FUNCTION_BLOCK StartStopEvent (* Basic Function Block Type *)
  (* Standard: 61499-2 *)
  (* Version 0.0, 10/21/2026, Schneider Electric, Template *)
  PACKAGE SE.Nereda;
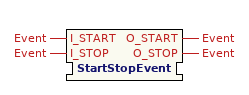
  EVENT_INPUT
    I_START; (* Normal Execution Request *)
    I_STOP;
  END_EVENT
  EVENT_OUTPUT
    O_START; (* Execution Confirmation *)
    O_STOP; (* Initialization Confirm *)
  END_EVENT
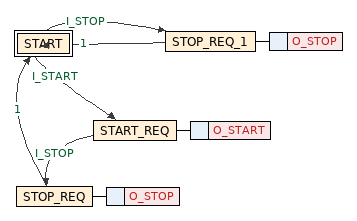
  EC_STATES
    START; (* Initial State *)
    START_REQ : -> O_START;
    STOP_REQ : -> O_STOP;
    STOP_REQ_1 : -> O_STOP;
  END_STATES
  EC_TRANSITIONS
    START TO START_REQ := I_START;
    START_REQ TO STOP_REQ := I_STOP;
    STOP_REQ TO START := 1;
    START TO STOP_REQ_1 := I_STOP;
    STOP_REQ_1 TO START := 1;
  END_TRANSITIONS
  ALGORITHM INIT IN ST: (* Initialization algorithm *)
;
  END_ALGORITHM
  ALGORITHM REQ IN ST: (* Normally executed algorithm *)
;
  END_ALGORITHM
END_FUNCTION_BLOCK
